Fanuc KAREL source: KD00001.KL

PROGRAM KD00001
%NOLOCKGROUP
%ALPHABETIZE
VAR
  I: INTEGER
  J: INTEGER
  B: BOOLEAN
  R: REAL
  S: STRING[80]
BEGIN
  I = 1
END KD00001
